(* IEC 61131-3 sources: llm-plc-st-eval/data/definitivo/gpt-4o-2024-08-06/B7/zero_shot, 3 files *)

(* ---- ejec_2.st ---- *)
Aquí tienes el código en Structured Text (ST) para la lógica de selección de la fuente de mando de una bomba, utilizando un FUNCTION_BLOCK llamado `SelBomba`. Este bloque de función recibe las entradas `modoAuto`, `btnManual` y `nivelBajo`, y entrega el estado de la bomba a través de la salida `bomba`.

```pascal
FUNCTION_BLOCK SelBomba
VAR_INPUT
    modoAuto : BOOL;    // Indica si el modo automático está activo
    btnManual : BOOL;   // Estado del botón manual
    nivelBajo : BOOL;   // Indica si el nivel bajo está activo
END_VAR

VAR_OUTPUT
    bomba : BOOL;       // Estado de la bomba
END_VAR

// Lógica de control de la bomba
// Si modo automático está activo, la bomba se enciende si nivelBajo está activo
// Si modo automático no está activo, la bomba sigue el estado del botón manual
bomba := (modoAuto AND nivelBajo) OR (NOT modoAuto AND btnManual);

END_FUNCTION_BLOCK
```

Este bloque de función `SelBomba` evalúa las condiciones de las entradas en cada ciclo de ejecución y determina el estado de la bomba en función del modo de operación seleccionado.

(* ---- ejec_3.st ---- *)
Aquí tienes el código en Structured Text (ST) para un FUNCTION_BLOCK llamado `SelBomba`, que implementa la lógica de selección de la fuente de mando de una bomba conforme a tu descripción:

```pascal
FUNCTION_BLOCK SelBomba
VAR_INPUT
    modoAuto : BOOL;    // Indica si el modo automático está activo
    btnManual : BOOL;   // Estado del botón manual
    nivelBajo : BOOL;   // Indica si el nivel bajo está activo
END_VAR
VAR_OUTPUT
    bomba : BOOL;       // Estado de la bomba
END_VAR

// Lógica de control de la bomba
bomba := (modoAuto AND nivelBajo) OR (NOT modoAuto AND btnManual);

END_FUNCTION_BLOCK
```

### Explicación:
- **modoAuto**: Entrada booleana que indica si el modo automático está activo.
- **btnManual**: Entrada booleana que representa el estado del botón manual.
- **nivelBajo**: Entrada booleana que indica si el nivel bajo está activo.
- **bomba**: Salida booleana que representa el estado de la bomba.

La lógica implementada en el bloque `SelBomba` establece que la bomba se enciende si:
- El modo automático está activo y el nivel bajo está activo, o
- El modo manual está activo (modo automático no activo) y el botón manual está presionado.

(* ---- ejec_1.st ---- *)
```pascal
PROGRAM SelBomba
VAR
    modoAuto : BOOL;    // Entrada: selecciona el modo automático
    btnManual : BOOL;   // Entrada: botón manual para encender la bomba
    nivelBajo : BOOL;   // Entrada: indica si el nivel es bajo
    bomba : BOOL;       // Salida: estado de la bomba
END_VAR

// Lógica de selección de la fuente de mando de la bomba
IF modoAuto THEN
    // Modo automático: la bomba se enciende si nivelBajo está activo
    bomba := nivelBajo;
ELSE
    // Modo manual: la bomba sigue el estado del botón manual
    bomba := btnManual;
END_IF;
```

Este código define un programa (`PROGRAM`) llamado `SelBomba` que implementa la lógica de control de una bomba basada en el modo de operación seleccionado (automático o manual). Las entradas son `modoAuto`, `btnManual` y `nivelBajo`, y la salida es `bomba`, que indica el estado actual de la bomba.
